FUNCTION_BLOCK FB_NCIMeina2_2000x1000 EXTENDS FB_RecipeBase

METHOD Build : BOOL
VAR
      i          : INT;
	  sRecipeName : STRING(255) := '\Hard Disk\Meina2_2000x1000.nc';
END_VAR

VAR_INST
    nBuildStep : INT;
    machineConfig : ST_GantryXYZ_Config;
END_VAR
Build := FALSE;

CASE nBuildStep OF
    0:
        _Busy := TRUE;
        _Done := FALSE;
        _Error := FALSE;
        
        _Config.GCodePath := sRecipeName; 
        
        ADSLOGSTR(ADSLOG_MSGTYPE_HINT, CONCAT('Builder: Skonfigurowano gotowy plik G-Code: ', sRecipeName), '');
        
        nBuildStep := 1000;

    1000:
        _Busy := FALSE;
        _Done := TRUE; 
        nBuildStep := 0;
        Build := TRUE;
        
END_CASE
END_METHOD

PROPERTY ExecutionRoute : E_ExecutionRoute
GET
ExecutionRoute := E_ExecutionRoute.eGCode;
END_GET
END_PROPERTY

END_FUNCTION_BLOCK

(* stored: Version 1.1.0.1, ProductVersion 3.1.4024.15
   POU FB_NCIMeina2_2000x1000: Id {22b8006b-85a6-4b7f-b0ea-19ab060d1e2b}, SpecialFunc None
   Method Build: Id {fa0b89f6-ef30-4f8b-ba6b-e1f90d3f2882}
   Property ExecutionRoute: Id {2522e725-4c9d-4aa7-9745-528a8d6a0bfc}
   Get Get: Id {c3e2079d-c741-4220-a7e8-afb21e7ed919} *)
